FUNCTION_BLOCK FB_StationPickup EXTENDS FB_RollerConveyor
// =============================================================
// STACJA ODBIORU - 13 (stosy dobre) I 16 (palety odrzucone)
// =============================================================
//
// Koniec drogi: ladunek stoi na czujnikach i zabiera go operator.
// Nie ma nastepnika, wiec zwolnienie miejsca musi wykryc sama
// stacja.
//
// Dwa sposoby, przelaczane nastawa Cfg.xPickupByButton:
//
//   TRUE  - operator potwierdza przyciskiem. Sprawdzamy wtedy,
//           czy ladunek faktycznie zniknal z czujnikow. Jesli
//           nie zniknal, nie robimy nic - przycisk nie jest
//           dowodem na to, ze cos zostalo zabrane.
//
//   FALSE - miejsce uznajemy za wolne po Cfg.tPickupTimeout
//           od zniknieca ladunku z czujnikow.
VAR_INPUT

	// Przycisk operatora "zabralem"
	xPickupButton	: BOOL;

END_VAR
VAR_OUTPUT

	// Czeka na odbior
	xWaitingPickup	: BOOL;

END_VAR
VAR

	tonPickup	: TON;
	rtrgButton	: R_TRIG;

END_VAR

SUPER^();

M_PickupCycle();

METHOD PROTECTED M_PickupCycle
VAR
	xFree	: BOOL;
END_VAR
xWaitingPickup := FALSE;

IF pP = 0 THEN
	RETURN;
END_IF

IF NOT pP^.Mem.xLoadPresent THEN
	tonPickup(IN := FALSE);
	rtrgButton(CLK := xPickupButton);
	RETURN;
END_IF

xWaitingPickup	:= TRUE;
eWait			:= WAIT_PICKUP;


// Pole czujnikow wolne. Przy wylaczonych czujnikach nie mamy
// czym tego stwierdzic - wtedy decyduje sam przycisk.
IF xSensUsable THEN
	xFree := xSensLoadNone;
ELSE
	xFree := TRUE;
END_IF


// --- potwierdzenie przyciskiem ---
IF pP^.Cfg.xPickupByButton THEN

	rtrgButton(CLK := xPickupButton);

	IF NOT rtrgButton.Q THEN
		RETURN;
	END_IF

	// Przycisk wcisniety, ale ladunek dalej lezy - nic nie robimy
	IF NOT xFree THEN
		RETURN;
	END_IF

	M_ClearLoad();
	RETURN;

END_IF


// --- odliczanie od zniknieca z czujnikow ---
rtrgButton(CLK := xPickupButton);

tonPickup(IN := xFree, PT := pP^.Cfg.tPickupTimeout);

IF tonPickup.Q THEN
	tonPickup(IN := FALSE);
	M_ClearLoad();
END_IF
END_METHOD

METHOD PROTECTED M_OperationRequired : BOOL
// Nie ma operacji technologicznej - ladunek po prostu czeka.
M_OperationRequired := FALSE;
END_METHOD

END_FUNCTION_BLOCK

(* stored: Version 1.1.0.1
   POU FB_StationPickup: Id {7b2d0a00-0000-4000-9000-000000000a00}, SpecialFunc None
   Method M_PickupCycle: Id {7b2d0a01-0000-4000-9000-000000000a01}
   Method M_OperationRequired: Id {7b2d0a02-0000-4000-9000-000000000a02} *)
